// TIA Portal V20 export
Screen "200RB04_V23"  1276x673
  ScreenItem "Graphic view_1" at 85,86 size 878x526  Type=HmiGraphicView
  ScreenItem "Line_Header_X0_Y64" at 0,64 size 1276x0  Type=HmiLine
  ScreenItem "permanentareaborderrectangle" at 0,0 size 0x0  Type=HmiRectangle
  ScreenItem "Button_Back" at 2,2 size 90x60  Type=HmiButton
  ScreenItem "Rectangle_3" at 0,0 size 166x43  Type=HmiRectangle
  ScreenItem "文本域_3" at 2,1 size 134x40  Type=HmiTextBox
  ScreenItem "圆_3" at 0,0 size 100x30  Type=HmiCircle
  ScreenItem "圆_4" at 0,0 size 100x30  Type=HmiCircle
  ScreenItem "文本域_9" at 963,181 size 134x40  Type=HmiTextBox
  ScreenItem "Line_7" at 552,324 size 18x141  Type=HmiLine
  ScreenItem "文本域_2" at 169,196 size 134x40  Type=HmiTextBox
  ScreenItem "文本域_4" at 437,85 size 134x40  Type=HmiTextBox
  ScreenItem "Rectangle_5" at 0,0 size 166x43  Type=HmiRectangle
  ScreenItem "文本域_5" at 2,1 size 134x40  Type=HmiTextBox
  ScreenItem "圆_1" at 0,0 size 100x30  Type=HmiCircle
  ScreenItem "圆_2" at 0,0 size 100x30  Type=HmiCircle
  ScreenItem "文本域_6" at 484,463 size 134x40  Type=HmiTextBox
  ScreenItem "Rectangle_13" at 0,0 size 166x43  Type=HmiRectangle
  ScreenItem "文本域_14" at 2,1 size 134x40  Type=HmiTextBox
  ScreenItem "圆_5" at 0,0 size 100x30  Type=HmiCircle
  ScreenItem "圆_6" at 0,0 size 100x30  Type=HmiCircle
  ScreenItem "文本域_1" at 618,560 size 134x40  Type=HmiTextBox
  ScreenItem "文本域_7" at 963,75 size 134x40  Type=HmiTextBox
  ScreenItem "文本域_8" at 213,98 size 134x40  Type=HmiTextBox
  ScreenItem "Title_ScreenOverview_X390_Y2_20" at 254,162 size 25x21  Type=HmiTextBox
  ScreenItem "Title_ScreenOverview_X390_Y2_21" at 281,162 size 25x21  Type=HmiTextBox
  ScreenItem "Title_ScreenOverview_X390_Y2_22" at 254,142 size 52x19  Type=HmiTextBox
  ScreenItem "Line_1" at 674,458 size 1x101  Type=HmiLine
  ScreenItem "Line_2" at 668,315 size 305x144  Type=HmiLine
  ScreenItem "Line_3" at 385,320 size 153x141  Type=HmiLine
  ScreenItem "Line_4" at 346,123 size 130x116  Type=HmiLine
  ScreenItem "Line_5" at 828,328 size 145x68  Type=HmiLine
  ScreenItem "Line_6" at 571,104 size 63x96  Type=HmiLine
  ScreenItem "Line_8" at 897,324 size 77x1  Type=HmiLine
  ScreenItem "Line_9" at 753,93 size 209x102  Type=HmiLine
  ScreenItem "Line_10" at 302,215 size 109x70  Type=HmiLine
  ScreenItem "Line_11" at 791,206 size 174x108  Type=HmiLine
  ScreenItem "Rectangle_10" at 0,0 size 52x43  Type=HmiRectangle
  ScreenItem "Title_ScreenOverview_X390_Y2_111" at 0,21 size 25x21  Type=HmiTextBox
  ScreenItem "Title_ScreenOverview_X390_Y2_90" at 27,21 size 25x21  Type=HmiTextBox
  ScreenItem "Title_ScreenOverview_X390_Y2_88" at 0,1 size 52x19  Type=HmiTextBox
  ScreenItem "Rectangle_9" at 525,505 size 52x43  Type=HmiRectangle
  ScreenItem "Title_ScreenOverview_X390_Y2_17" at 525,526 size 25x21  Type=HmiTextBox
  ScreenItem "Title_ScreenOverview_X390_Y2_18" at 552,526 size 25x21  Type=HmiTextBox
  ScreenItem "Title_ScreenOverview_X390_Y2_19" at 525,506 size 52x19  Type=HmiTextBox
  ScreenItem "Title_ScreenOverview_X390_Y2_11" at 210,260 size 25x21  Type=HmiTextBox
  ScreenItem "Title_ScreenOverview_X390_Y2_12" at 237,260 size 25x21  Type=HmiTextBox
  ScreenItem "Title_ScreenOverview_X390_Y2_13" at 210,240 size 52x19  Type=HmiTextBox
  ScreenItem "Title_ScreenOverview_X390_Y2_5" at 478,149 size 25x21  Type=HmiTextBox
  ScreenItem "Title_ScreenOverview_X390_Y2_6" at 505,149 size 25x21  Type=HmiTextBox
  ScreenItem "Title_ScreenOverview_X390_Y2_7" at 478,129 size 52x19  Type=HmiTextBox
  ScreenItem "Title_ScreenOverview_X390_Y2_23" at 659,622 size 25x21  Type=HmiTextBox
  ScreenItem "Title_ScreenOverview_X390_Y2_24" at 686,622 size 25x21  Type=HmiTextBox
  ScreenItem "Title_ScreenOverview_X390_Y2_25" at 659,602 size 52x19  Type=HmiTextBox
  ScreenItem "Title_ScreenOverview_X390_Y2_26" at 1004,138 size 25x21  Type=HmiTextBox
  ScreenItem "Title_ScreenOverview_X390_Y2_27" at 1031,138 size 25x21  Type=HmiTextBox
  ScreenItem "Title_ScreenOverview_X390_Y2_28" at 1004,118 size 52x19  Type=HmiTextBox
  ScreenItem "Title_ScreenOverview_X390_Y2_2" at 392,4 size 510x57  Type=HmiTextBox
  ScreenItem "Title_ScreenOverview_X390_Y2_1" at 1130,78 size 139x57  Type=HmiTextBox
  ScreenItem "Title_ScreenOverview_X390_Y2_3" at 1130,144 size 139x57  Type=HmiTextBox
  ScreenItem "Title_ScreenOverview_X390_Y2_4" at 1130,144 size 139x57  Type=HmiTextBox
  ScreenItem "Rectangle_6" at 210,239 size 52x43  Type=HmiRectangle
  ScreenItem "Rectangle_2" at 478,128 size 52x43  Type=HmiRectangle
  ScreenItem "Rectangle_1" at 659,601 size 52x43  Type=HmiRectangle
  ScreenItem "Rectangle_12" at 1004,116 size 52x43  Type=HmiRectangle
  ScreenItem "Rectangle_8" at 254,141 size 52x43  Type=HmiRectangle
  ScreenItem "Rectangle_4" at 0,0 size 166x43  Type=HmiRectangle
  ScreenItem "文本域_10" at 2,1 size 134x40  Type=HmiTextBox
  ScreenItem "圆_7" at 0,0 size 100x30  Type=HmiCircle
  ScreenItem "圆_8" at 0,0 size 100x30  Type=HmiCircle
  ScreenItem "Fusszeile_Button_ManualOPMode1_1" at 1179,3 size 90x60  Type=HmiButton
